TYPE ET_MC_ControllerMode :
(
	ET_MC_ControllerMode_eCMUndefined,
	ET_MC_ControllerMode_eCMTorque,
	ET_MC_ControllerMode_eCMVelocity,
	ET_MC_ControllerMode_eCMPosition,
	ET_MC_ControllerMode_eCMCurrent
	
);
END_TYPE

(* stored: Version 1.1.0.1, ProductVersion 3.1.4024.15
   DUT ET_MC_ControllerMode: Id {dbe08c0f-cb10-44fd-9f5e-1d40fadfe6dd} *)
